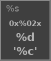
VISUALIZATION FRM_Segment  // 51x61
VAR_IN_OUT
   nValue: USINT;
END_VAR
VAR_INPUT
   nIndex: USINT;  
END_VAR
    Rectangle (0,0 51x61)
    Textfield (10,18 31x11), "0x%02x", text variable: nValue
    Textfield (3,3 21x11), "%s", text variable: TO_STRING(nIndex)
    Textfield (10,32 31x11), "%d", text variable: nValue
    Textfield (0,46 51x11), "'%c'", text variable: nValue, invisible if: (nValue < 32) OR (nValue > 126)
END_VISUALIZATION

(* stored: Version 1.1.0.1
   Visu FRM_Segment: Id {7078dc8b-64bc-0fc6-3a8b-7aed92bcd66f} *)
